# EPICS autosave request: 1.5.0/debian-12/7.0.10/modules/motor-4b22ac9/db/pseudoMotor_settings.req
# FILE... pseudoMotor_settings.req
$(P)$(M).DHLM
$(P)$(M).DLLM
$(P)$(M).TWV
$(P)$(M).DISA
$(P)$(M).DISP
$(P)$(M).OFF
$(P)$(M).VELO
$(P)$(M)C1
$(P)$(M)C2
$(P)$(M)C3
$(P)$(M)C4
$(P)$(M)C5
$(P)$(M)_able.VAL
